// TIA Portal V20 export
DATA_BLOCK "T6_Datos"   // DB43900
{ S7_Optimized_Access := 'TRUE' }
AUTHOR : IA
FAMILY : PRUEBA
VERSION : 0.1
// Tanda 2: datos
// stored: AutoNumber false
   VAR
      Dtl_1 : DTL;
      Dtl_2 : DTL;
      Dtl_3 : DTL;
      Dtl_Ahora : DTL;
      T_1500ms : Time := T#1500MS;
      T_Out : Time;
      DI_Out : DInt;
      DInt_2000 : DInt := 2000;
      T_1h : Time := T#1H;
      Fecha : Date := D#2026-03-04;
      Hora : Time_Of_Day := TOD#12:30:00;
      Ret_Leer : Int;
      Ret_Escribir : Int;
      Falso : Bool := false;
      S_ABCDEF : String := 'ABCDEF';
      S_Out : String;
      Int_123 : Int := 123;
      S_456 : String := '456';
      Int_3 : Int := 3;
      Int_2 : Int := 2;
      Int_2b : Int := 2;
      Int_1 : Int := 1;
      Int_3b : Int := 3;
      S_ABEF : String := 'ABEF';
      S_CD : String := 'CD';
      S_XY : String := 'XY';
      S_1A2B : String := '1A2B';
      Int_4 : Int := 4;
      UInt_2 : UInt := 2;
      Bytes : Array[0..9] of Byte;
      W_Ret : Word;
      Char_A : Char := 'A';
      Char_A2 : Char := 'A';
      T_desde_DInt : Time;
      T_Diff : Time;
      D_Comb : DTL;
      WrLoc_Mem : Bool;
      Ret_WrLoc : Int := -1;
      WrSys_Mem : Bool;
      Ret_WrSys : Int := -1;
      D_Sys : DTL;
      Dtl_1_Copia : DTL;
      S_desde_Int : String;
      Int_vuelta : Int;
      I_desde_S : Int;
      LEFT_Out : String;
      RIGHT_Out : String;
      MID_Out : String;
      DELETE_Out : String;
      INSERT_Out : String;
      REPLACE_Out : String;
      FIND_Out : Int;
      HTA_Out : String;
      W_Ret2 : Word;
      Bytes_HTA : Array[0..9] of Byte;
      Escrito_S : Bool;
   END_VAR
BEGIN
END_DATA_BLOCK
